(* Logix 5000 project; controller TFF vendor 1 type 14 code 107 rev 34.11; software revision 34.03; part 32 of 36 *)
(* tags used below, declared in another part *)
   FlowPathControl : FlowPathControl;   // Flow Path Control
   Options : Options;   // Options List
   PCV001_Control : PCV_Control;   // PCV001 Control UDT
   PCV101_Control : PCV_Control;   // PCV101 Control UDT
   PipeAnimation : PipeAnimation;   // HMI Pipe Animation Array
   XV001 : ALIAS FOR Valve[0];   // XV001
   XV002 : ALIAS FOR Valve[1];   // XV002
   XV004 : ALIAS FOR Valve[3];   // XV004
   XV005 : ALIAS FOR Valve[4];   // XV005
   XV006 : ALIAS FOR Valve[19];
   XV007 : ALIAS FOR Valve[20];
   XV102 : ALIAS FOR Valve[5];   // XV102
   XV401 : ALIAS FOR Valve[6];   // XV401
   XV402 : ALIAS FOR Valve[7];   // XV402
   XV403 : ALIAS FOR Valve[15];
   XV404 : ALIAS FOR Valve[16];
   XV405 : ALIAS FOR Valve[17];
   XV406 : ALIAS FOR Valve[18];
   XV411 : ALIAS FOR Valve[8];   // XV411
   XV421 : ALIAS FOR Valve[9];   // XV421
   XV431 : ALIAS FOR Valve[10];   // XV431
   XV441 : ALIAS FOR Valve[11];   // XV441
   XV501 : ALIAS FOR Valve[12];   // XV501
   XV502 : ALIAS FOR Valve[13];   // XV502
(* Process, continued *)

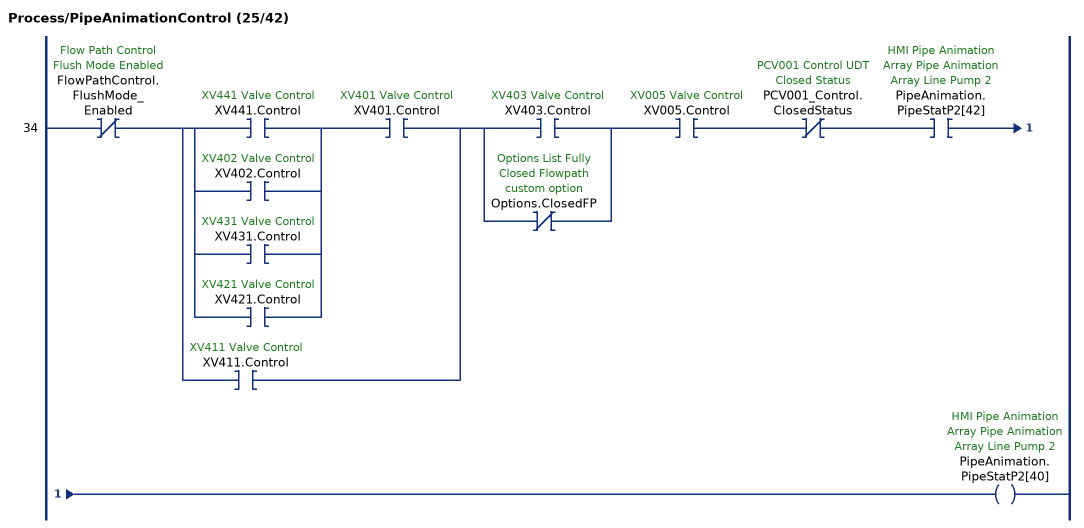
   [picture p389: Process/PipeAnimationControl rungs 34-34]
   34: XIO(FlowPathControl.FlushMode_Enabled)[[XIC(XV441.Control) ,XIC(XV402.Control) ,XIC(XV431.Control) ,XIC(XV421.Control) ] XIC(XV401.Control) ,XIC(XV411.Control) ][XIC(XV403.Control) ,XIO(Options.ClosedFP) ]XIC(XV005.Control)XIO(PCV001_Control.ClosedStatus)XIC(PipeAnimation.PipeStatP2[42])OTE(PipeAnimation.PipeStatP2[40]);
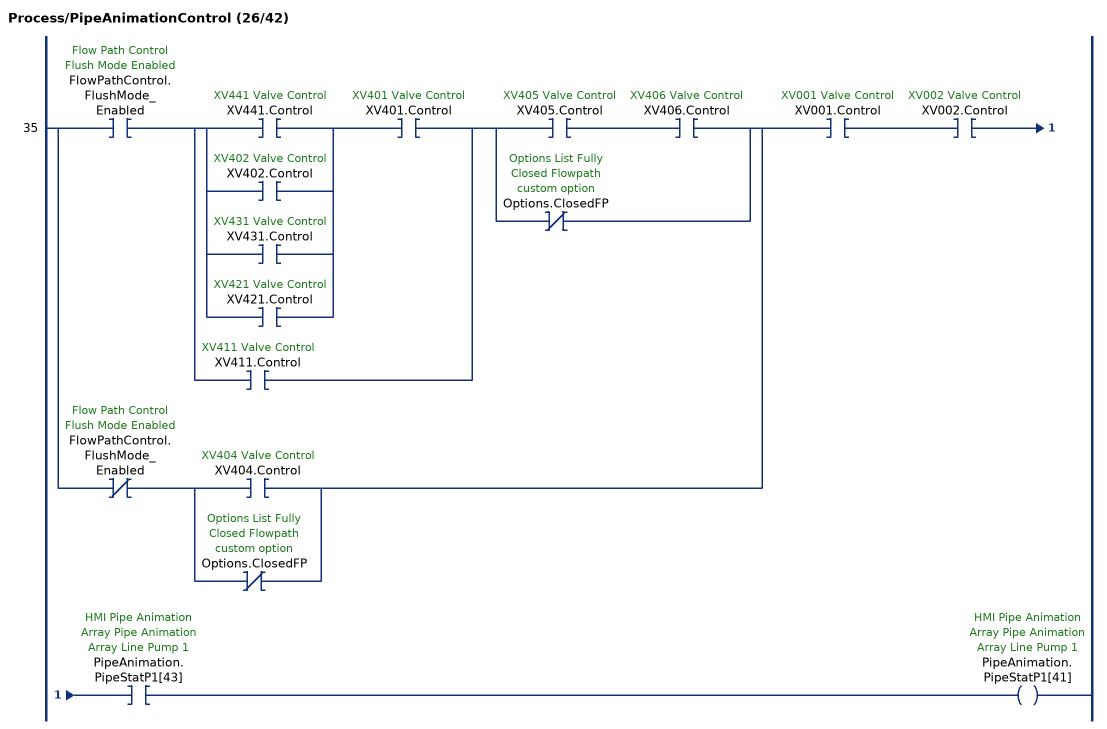
   35: [XIC(FlowPathControl.FlushMode_Enabled) [[XIC(XV441.Control) ,XIC(XV402.Control) ,XIC(XV431.Control) ,XIC(XV421.Control) ] XIC(XV401.Control) ,XIC(XV411.Control) ] [XIC(XV405.Control) XIC(XV406.Control) ,XIO(Options.ClosedFP) ] ,XIO(FlowPathControl.FlushMode_Enabled) [XIC(XV404.Control) ,XIO(Options.ClosedFP) ] ]XIC(XV001.Control)XIC(XV002.Control)XIC(PipeAnimation.PipeStatP1[43])OTE(PipeAnimation.PipeStatP1[41]);
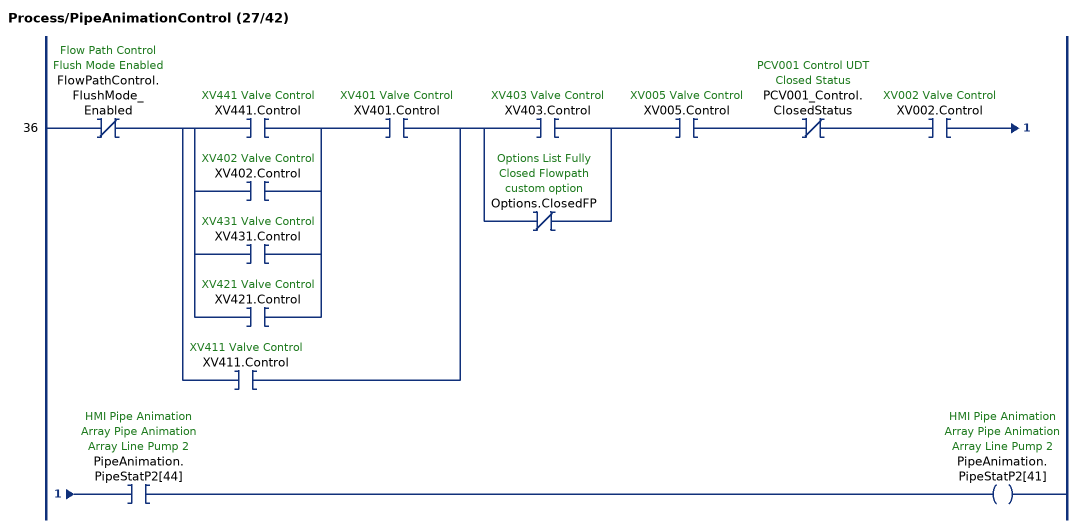
   36: XIO(FlowPathControl.FlushMode_Enabled)[[XIC(XV441.Control) ,XIC(XV402.Control) ,XIC(XV431.Control) ,XIC(XV421.Control) ] XIC(XV401.Control) ,XIC(XV411.Control) ][XIC(XV403.Control) ,XIO(Options.ClosedFP) ]XIC(XV005.Control)XIO(PCV001_Control.ClosedStatus)XIC(XV002.Control)XIC(PipeAnimation.PipeStatP2[44])OTE(PipeAnimation.PipeStatP2[41]);
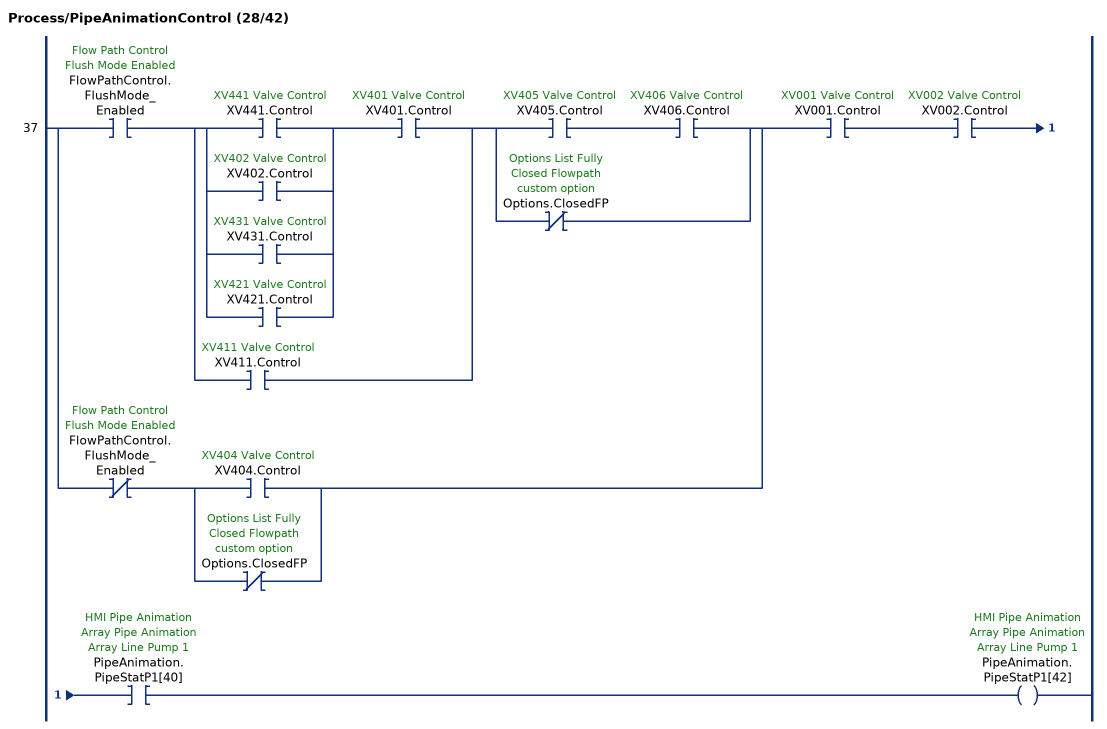
   37: [XIC(FlowPathControl.FlushMode_Enabled) [[XIC(XV441.Control) ,XIC(XV402.Control) ,XIC(XV431.Control) ,XIC(XV421.Control) ] XIC(XV401.Control) ,XIC(XV411.Control) ] [XIC(XV405.Control) XIC(XV406.Control) ,XIO(Options.ClosedFP) ] ,XIO(FlowPathControl.FlushMode_Enabled) [XIC(XV404.Control) ,XIO(Options.ClosedFP) ] ]XIC(XV001.Control)XIC(XV002.Control)XIC(PipeAnimation.PipeStatP1[40])OTE(PipeAnimation.PipeStatP1[42]);
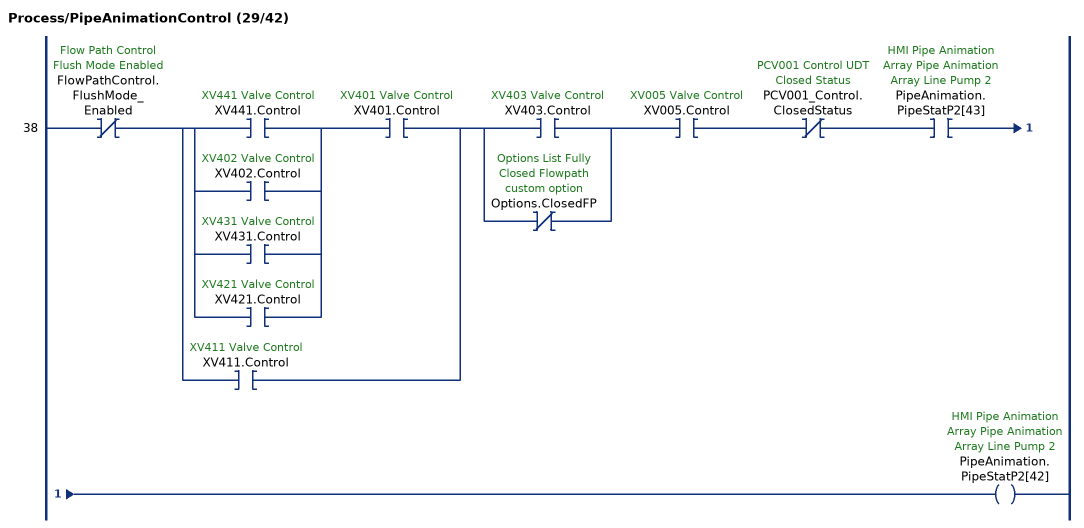
   38: XIO(FlowPathControl.FlushMode_Enabled)[[XIC(XV441.Control) ,XIC(XV402.Control) ,XIC(XV431.Control) ,XIC(XV421.Control) ] XIC(XV401.Control) ,XIC(XV411.Control) ][XIC(XV403.Control) ,XIO(Options.ClosedFP) ]XIC(XV005.Control)XIO(PCV001_Control.ClosedStatus)XIC(PipeAnimation.PipeStatP2[43])OTE(PipeAnimation.PipeStatP2[42]);
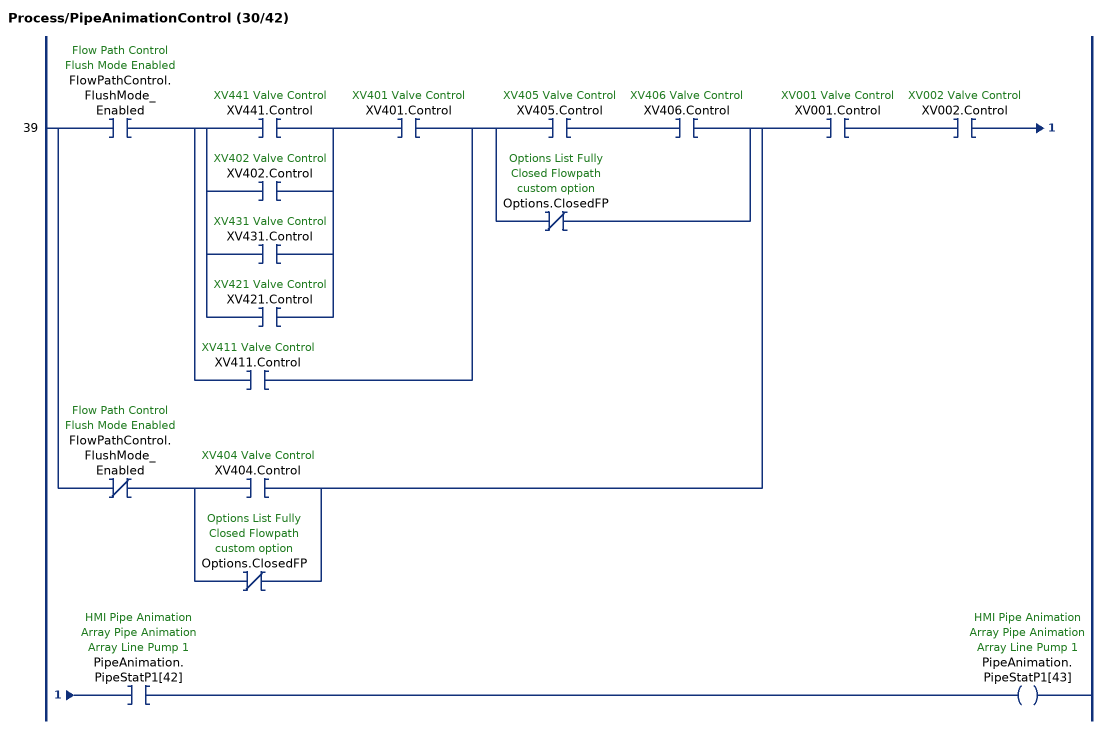
   39: [XIC(FlowPathControl.FlushMode_Enabled) [[XIC(XV441.Control) ,XIC(XV402.Control) ,XIC(XV431.Control) ,XIC(XV421.Control) ] XIC(XV401.Control) ,XIC(XV411.Control) ] [XIC(XV405.Control) XIC(XV406.Control) ,XIO(Options.ClosedFP) ] ,XIO(FlowPathControl.FlushMode_Enabled) [XIC(XV404.Control) ,XIO(Options.ClosedFP) ] ]XIC(XV001.Control)XIC(XV002.Control)XIC(PipeAnimation.PipeStatP1[42])OTE(PipeAnimation.PipeStatP1[43]);
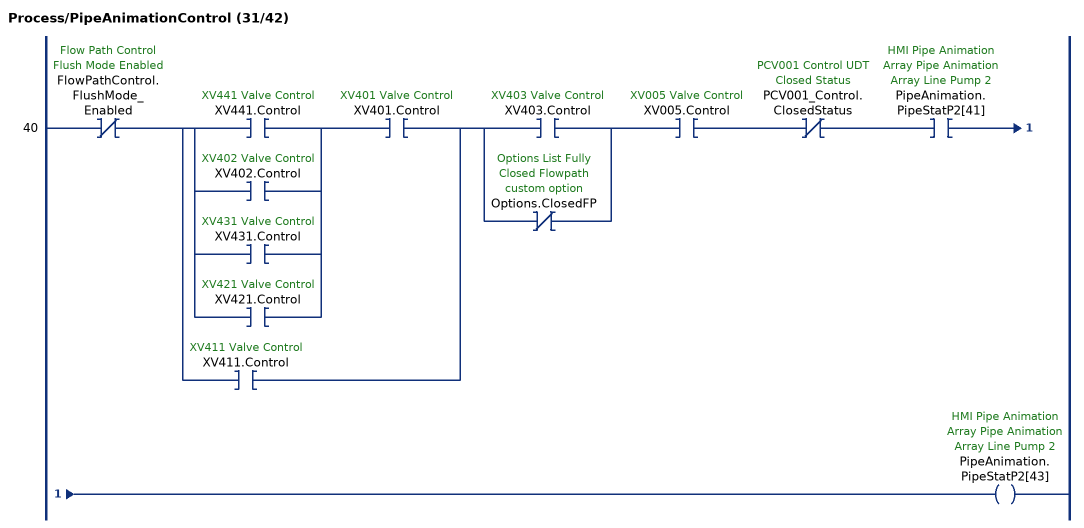
   40: XIO(FlowPathControl.FlushMode_Enabled)[[XIC(XV441.Control) ,XIC(XV402.Control) ,XIC(XV431.Control) ,XIC(XV421.Control) ] XIC(XV401.Control) ,XIC(XV411.Control) ][XIC(XV403.Control) ,XIO(Options.ClosedFP) ]XIC(XV005.Control)XIO(PCV001_Control.ClosedStatus)XIC(PipeAnimation.PipeStatP2[41])OTE(PipeAnimation.PipeStatP2[43]);
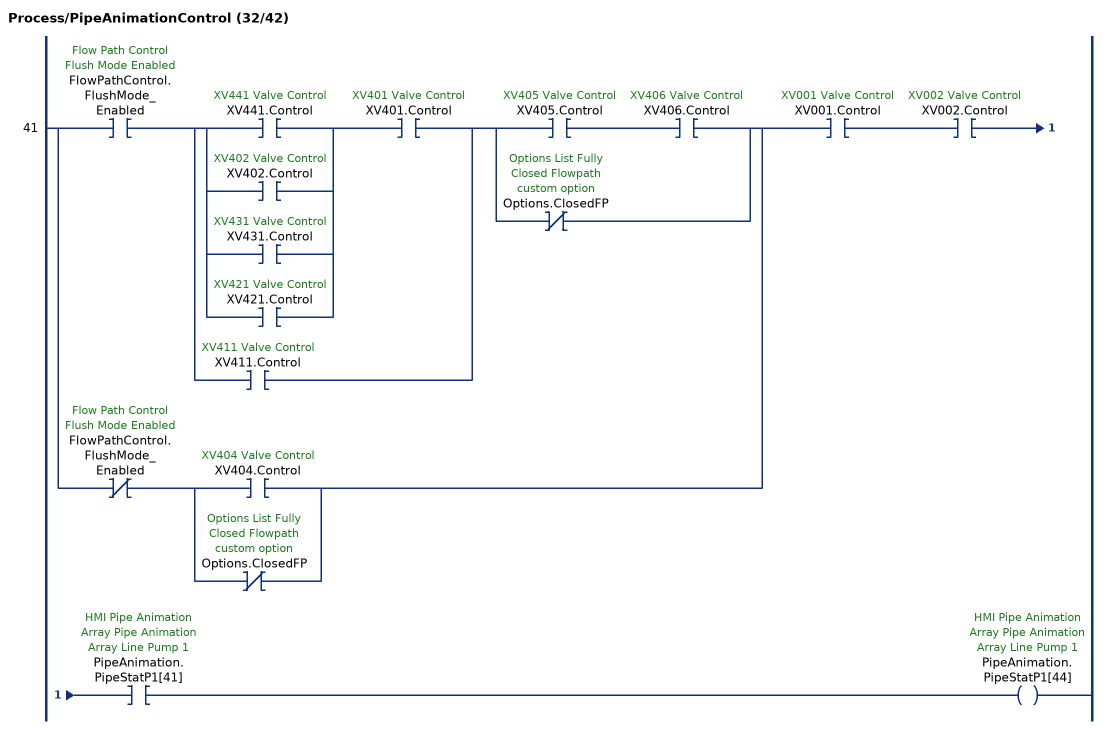
   41: [XIC(FlowPathControl.FlushMode_Enabled) [[XIC(XV441.Control) ,XIC(XV402.Control) ,XIC(XV431.Control) ,XIC(XV421.Control) ] XIC(XV401.Control) ,XIC(XV411.Control) ] [XIC(XV405.Control) XIC(XV406.Control) ,XIO(Options.ClosedFP) ] ,XIO(FlowPathControl.FlushMode_Enabled) [XIC(XV404.Control) ,XIO(Options.ClosedFP) ] ]XIC(XV001.Control)XIC(XV002.Control)XIC(PipeAnimation.PipeStatP1[41])OTE(PipeAnimation.PipeStatP1[44]);
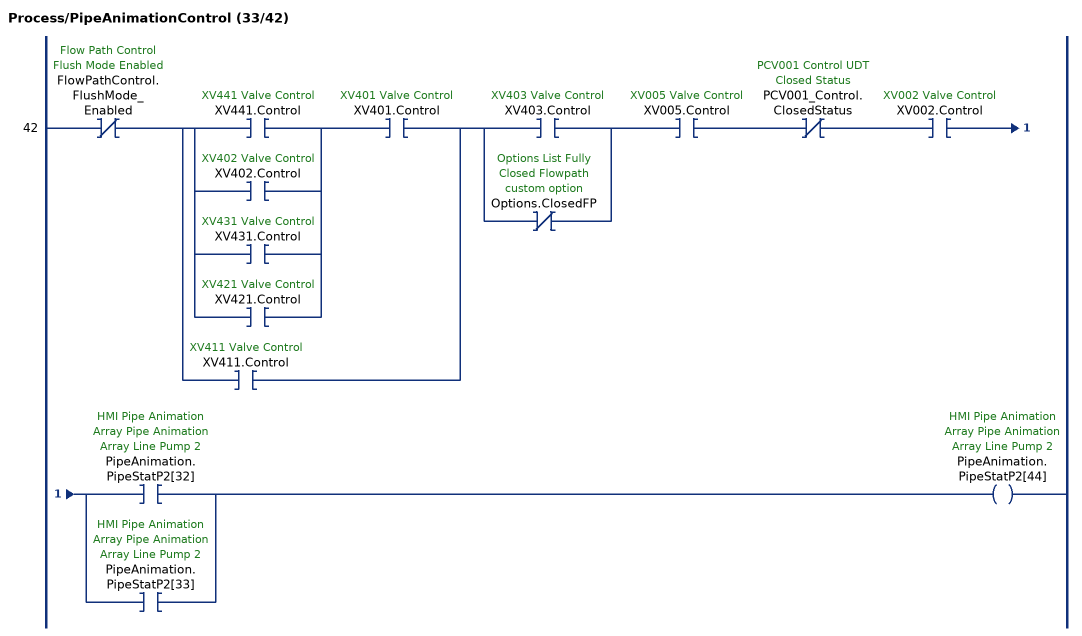
   42: XIO(FlowPathControl.FlushMode_Enabled)[[XIC(XV441.Control) ,XIC(XV402.Control) ,XIC(XV431.Control) ,XIC(XV421.Control) ] XIC(XV401.Control) ,XIC(XV411.Control) ][XIC(XV403.Control) ,XIO(Options.ClosedFP) ]XIC(XV005.Control)XIO(PCV001_Control.ClosedStatus)XIC(XV002.Control)[XIC(PipeAnimation.PipeStatP2[32]) ,XIC(PipeAnimation.PipeStatP2[33]) ]OTE(PipeAnimation.PipeStatP2[44]);
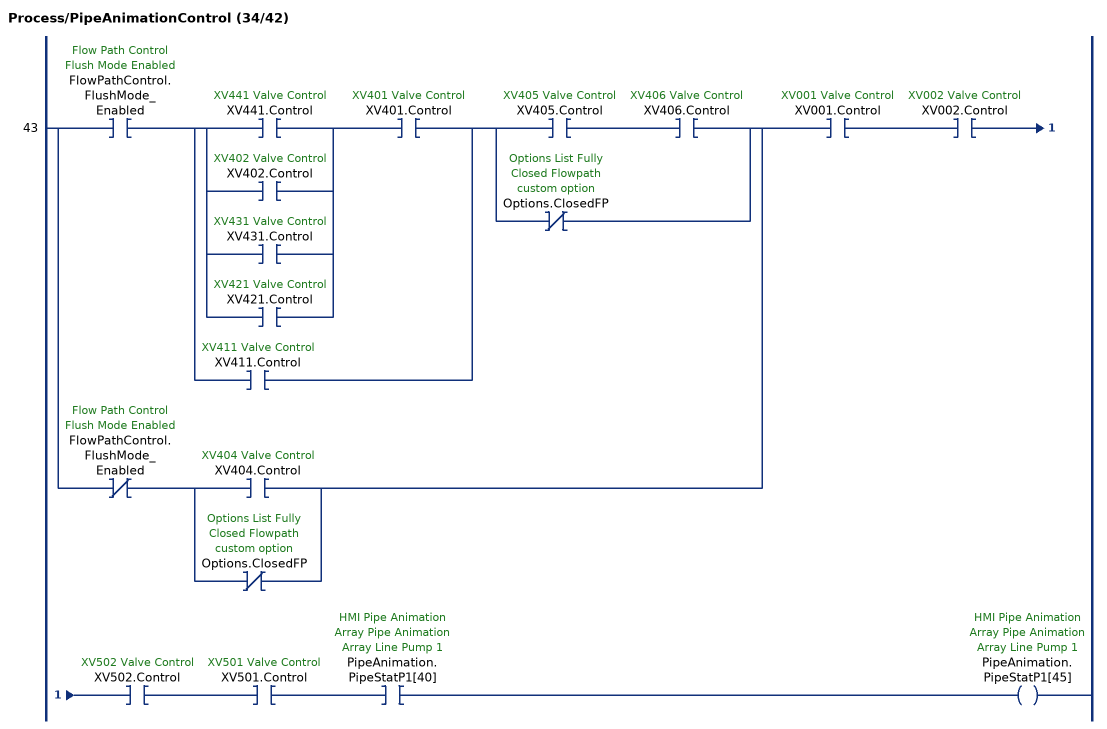
   43: [XIC(FlowPathControl.FlushMode_Enabled) [[XIC(XV441.Control) ,XIC(XV402.Control) ,XIC(XV431.Control) ,XIC(XV421.Control) ] XIC(XV401.Control) ,XIC(XV411.Control) ] [XIC(XV405.Control) XIC(XV406.Control) ,XIO(Options.ClosedFP) ] ,XIO(FlowPathControl.FlushMode_Enabled) [XIC(XV404.Control) ,XIO(Options.ClosedFP) ] ]XIC(XV001.Control)XIC(XV002.Control)XIC(XV502.Control)XIC(XV501.Control)XIC(PipeAnimation.PipeStatP1[40])OTE(PipeAnimation.PipeStatP1[45]);
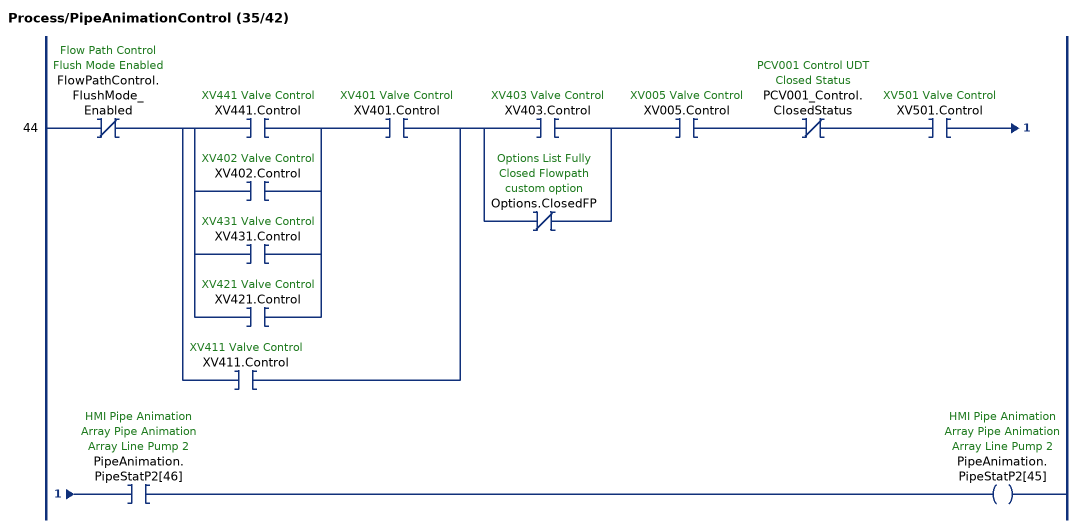
   44: XIO(FlowPathControl.FlushMode_Enabled)[[XIC(XV441.Control) ,XIC(XV402.Control) ,XIC(XV431.Control) ,XIC(XV421.Control) ] XIC(XV401.Control) ,XIC(XV411.Control) ][XIC(XV403.Control) ,XIO(Options.ClosedFP) ]XIC(XV005.Control)XIO(PCV001_Control.ClosedStatus)XIC(XV501.Control)XIC(PipeAnimation.PipeStatP2[46])OTE(PipeAnimation.PipeStatP2[45]);
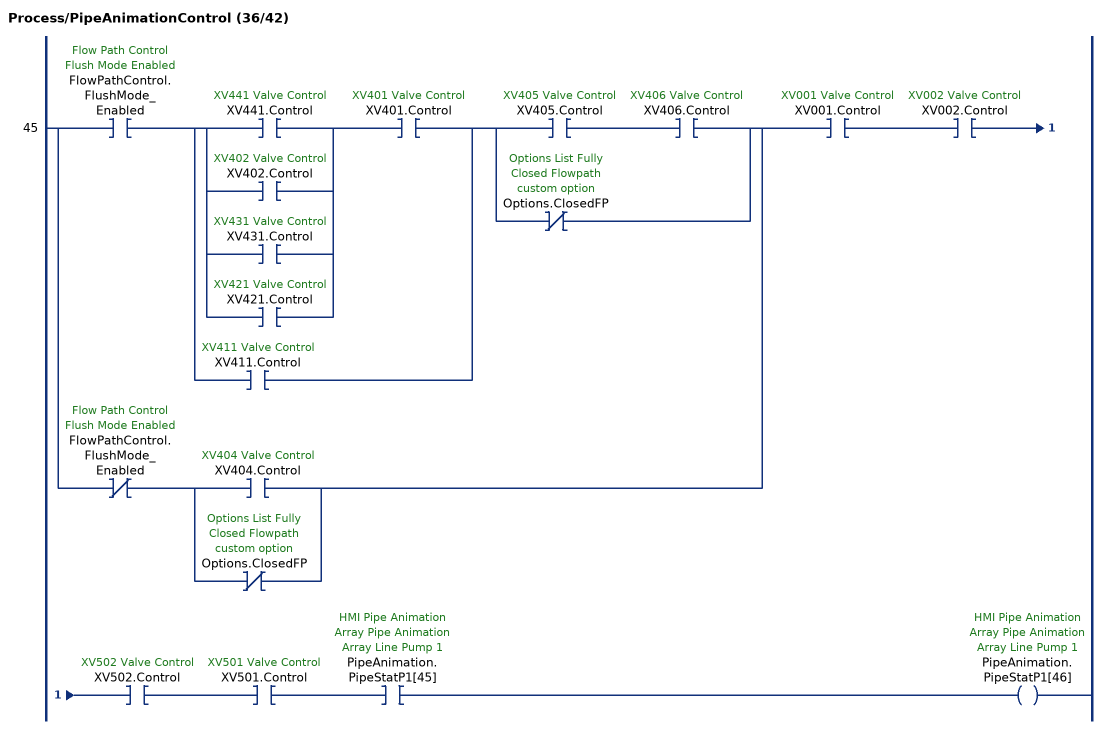
   45: [XIC(FlowPathControl.FlushMode_Enabled) [[XIC(XV441.Control) ,XIC(XV402.Control) ,XIC(XV431.Control) ,XIC(XV421.Control) ] XIC(XV401.Control) ,XIC(XV411.Control) ] [XIC(XV405.Control) XIC(XV406.Control) ,XIO(Options.ClosedFP) ] ,XIO(FlowPathControl.FlushMode_Enabled) [XIC(XV404.Control) ,XIO(Options.ClosedFP) ] ]XIC(XV001.Control)XIC(XV002.Control)XIC(XV502.Control)XIC(XV501.Control)XIC(PipeAnimation.PipeStatP1[45])OTE(PipeAnimation.PipeStatP1[46]);
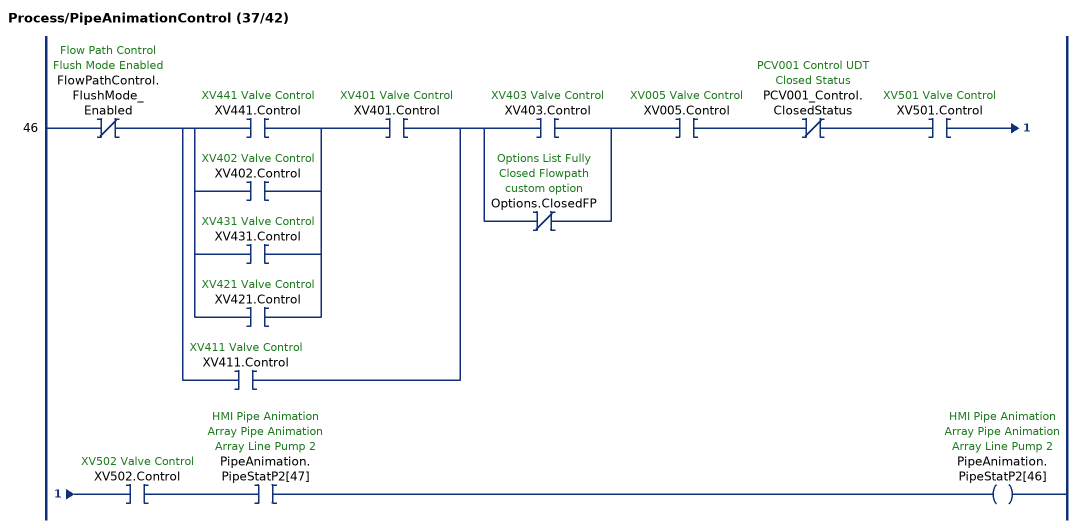
   46: XIO(FlowPathControl.FlushMode_Enabled)[[XIC(XV441.Control) ,XIC(XV402.Control) ,XIC(XV431.Control) ,XIC(XV421.Control) ] XIC(XV401.Control) ,XIC(XV411.Control) ][XIC(XV403.Control) ,XIO(Options.ClosedFP) ]XIC(XV005.Control)XIO(PCV001_Control.ClosedStatus)XIC(XV501.Control)XIC(XV502.Control)XIC(PipeAnimation.PipeStatP2[47])OTE(PipeAnimation.PipeStatP2[46]);
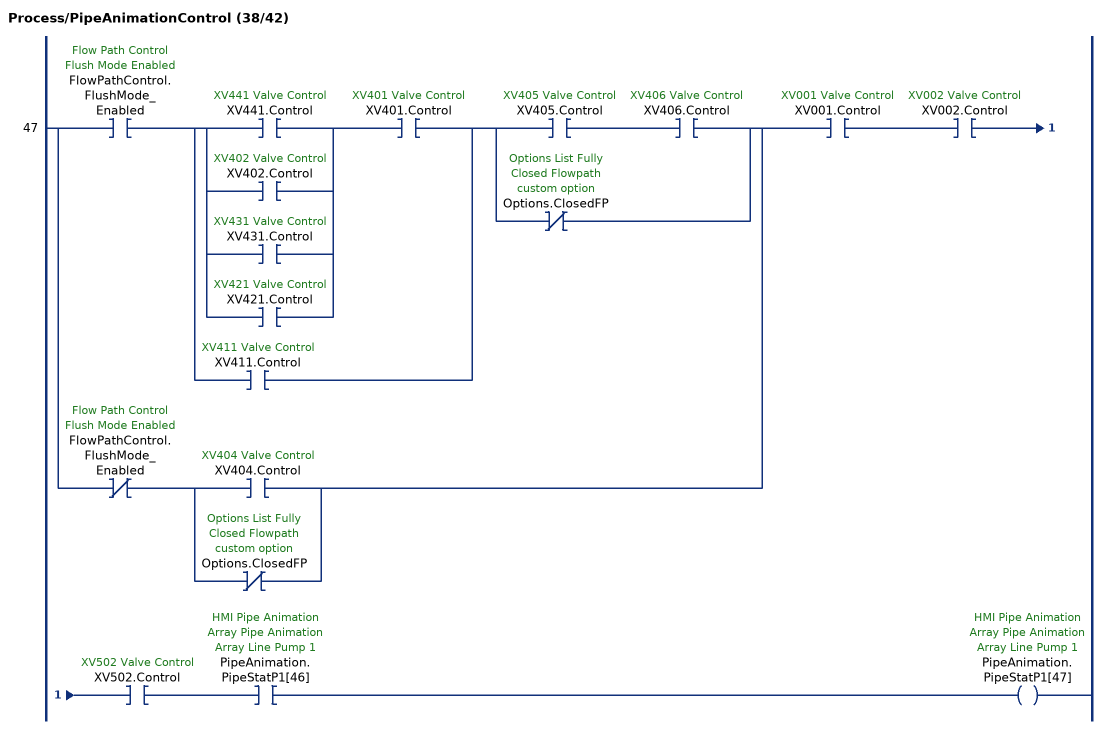
   47: [XIC(FlowPathControl.FlushMode_Enabled) [[XIC(XV441.Control) ,XIC(XV402.Control) ,XIC(XV431.Control) ,XIC(XV421.Control) ] XIC(XV401.Control) ,XIC(XV411.Control) ] [XIC(XV405.Control) XIC(XV406.Control) ,XIO(Options.ClosedFP) ] ,XIO(FlowPathControl.FlushMode_Enabled) [XIC(XV404.Control) ,XIO(Options.ClosedFP) ] ]XIC(XV001.Control)XIC(XV002.Control)XIC(XV502.Control)XIC(PipeAnimation.PipeStatP1[46])OTE(PipeAnimation.PipeStatP1[47]);
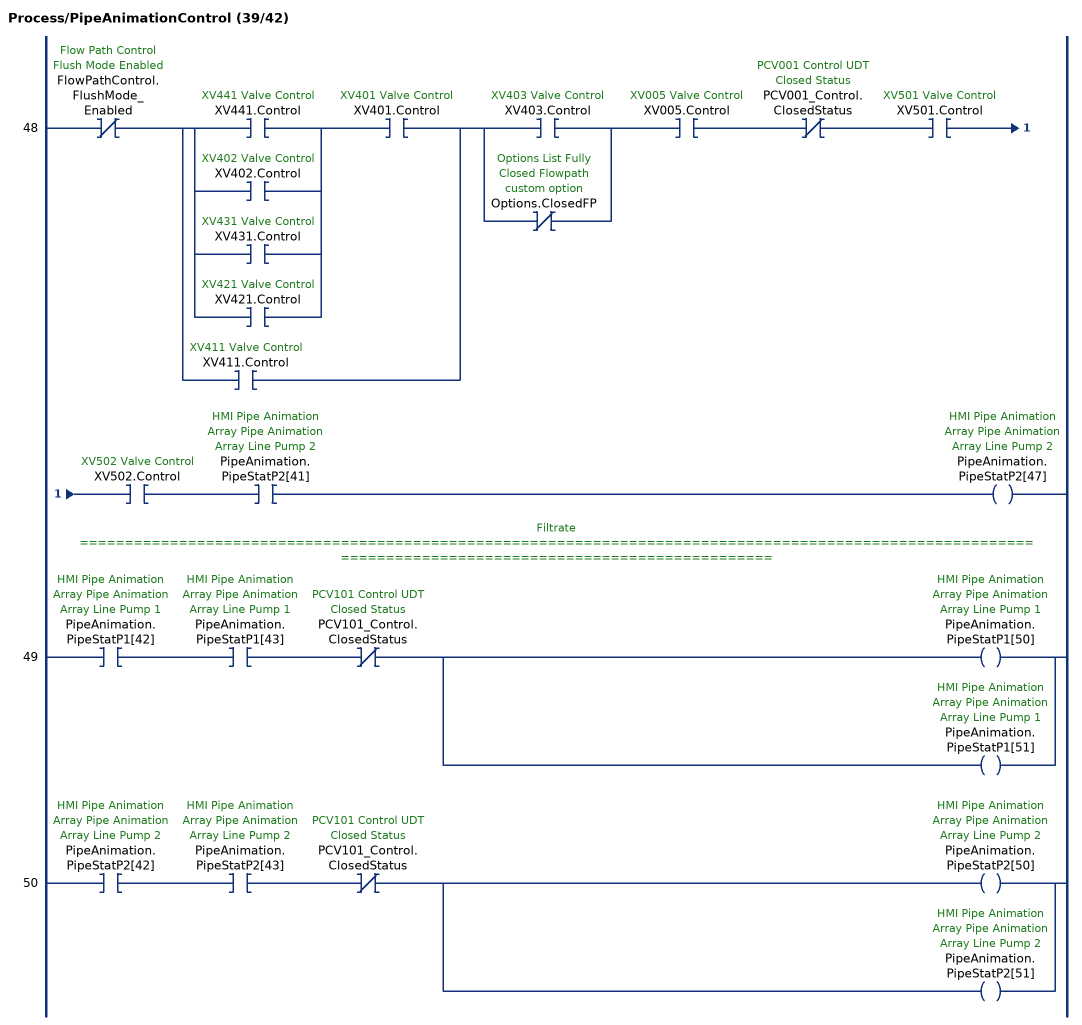
   48: XIO(FlowPathControl.FlushMode_Enabled)[[XIC(XV441.Control) ,XIC(XV402.Control) ,XIC(XV431.Control) ,XIC(XV421.Control) ] XIC(XV401.Control) ,XIC(XV411.Control) ][XIC(XV403.Control) ,XIO(Options.ClosedFP) ]XIC(XV005.Control)XIO(PCV001_Control.ClosedStatus)XIC(XV501.Control)XIC(XV502.Control)XIC(PipeAnimation.PipeStatP2[41])OTE(PipeAnimation.PipeStatP2[47]);
   // Filtrate
   // ==========================================================================================================================================================
   49: XIC(PipeAnimation.PipeStatP1[42])XIC(PipeAnimation.PipeStatP1[43])XIO(PCV101_Control.ClosedStatus)[OTE(PipeAnimation.PipeStatP1[50]) ,OTE(PipeAnimation.PipeStatP1[51]) ];
   50: XIC(PipeAnimation.PipeStatP2[42])XIC(PipeAnimation.PipeStatP2[43])XIO(PCV101_Control.ClosedStatus)[OTE(PipeAnimation.PipeStatP2[50]) ,OTE(PipeAnimation.PipeStatP2[51]) ];
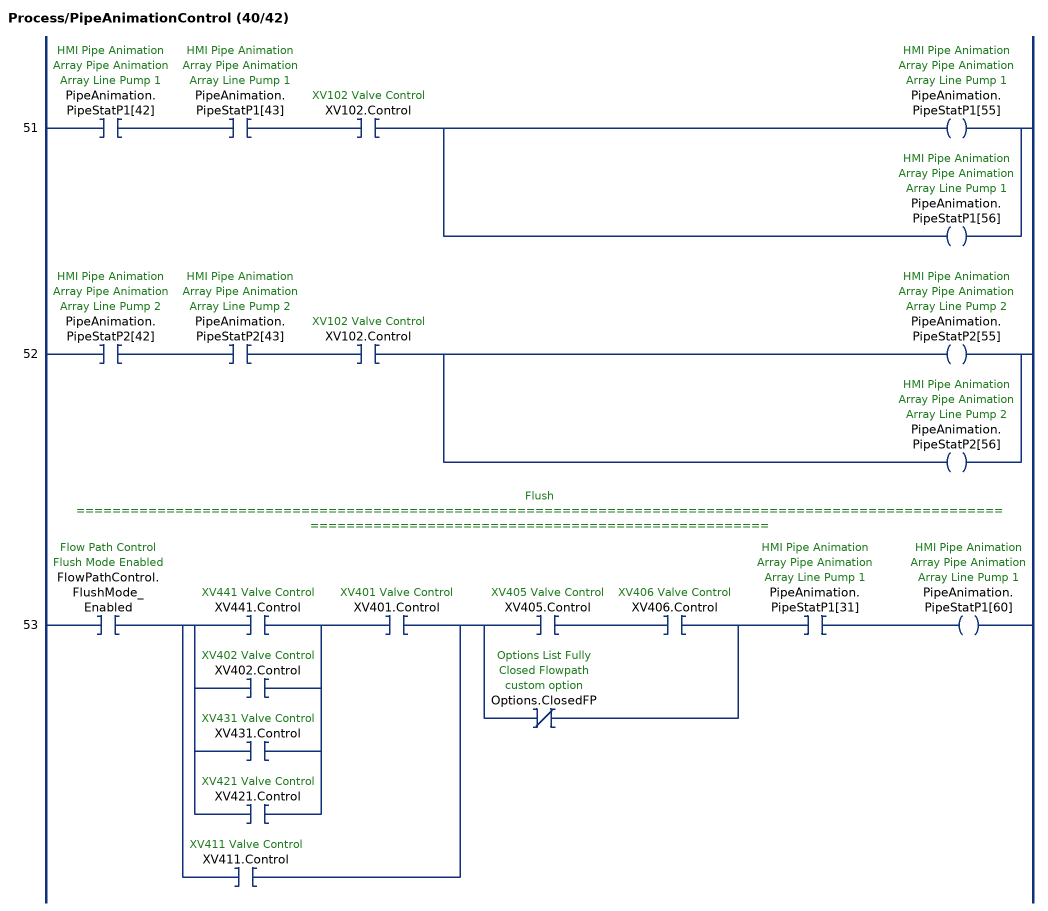
   51: XIC(PipeAnimation.PipeStatP1[42])XIC(PipeAnimation.PipeStatP1[43])XIC(XV102.Control)[OTE(PipeAnimation.PipeStatP1[55]) ,OTE(PipeAnimation.PipeStatP1[56]) ];
   52: XIC(PipeAnimation.PipeStatP2[42])XIC(PipeAnimation.PipeStatP2[43])XIC(XV102.Control)[OTE(PipeAnimation.PipeStatP2[55]) ,OTE(PipeAnimation.PipeStatP2[56]) ];
   // Flush
   // ==========================================================================================================================================================
   53: XIC(FlowPathControl.FlushMode_Enabled)[[XIC(XV441.Control) ,XIC(XV402.Control) ,XIC(XV431.Control) ,XIC(XV421.Control) ] XIC(XV401.Control) ,XIC(XV411.Control) ][XIC(XV405.Control) XIC(XV406.Control) ,XIO(Options.ClosedFP) ]XIC(PipeAnimation.PipeStatP1[31])OTE(PipeAnimation.PipeStatP1[60]);
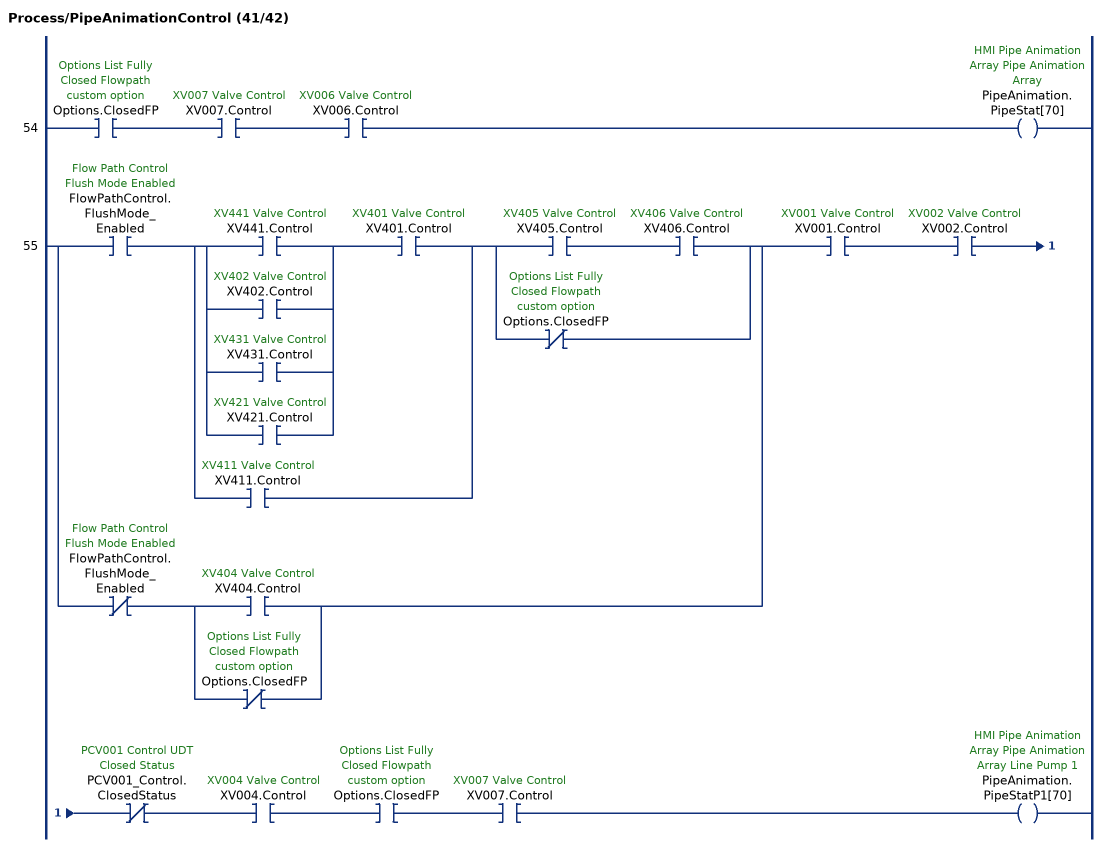
   54: XIC(Options.ClosedFP)XIC(XV007.Control)XIC(XV006.Control)OTE(PipeAnimation.PipeStat[70]);
   55: [XIC(FlowPathControl.FlushMode_Enabled) [[XIC(XV441.Control) ,XIC(XV402.Control) ,XIC(XV431.Control) ,XIC(XV421.Control) ] XIC(XV401.Control) ,XIC(XV411.Control) ] [XIC(XV405.Control) XIC(XV406.Control) ,XIO(Options.ClosedFP) ] ,XIO(FlowPathControl.FlushMode_Enabled) [XIC(XV404.Control) ,XIO(Options.ClosedFP) ] ]XIC(XV001.Control)XIC(XV002.Control)XIO(PCV001_Control.ClosedStatus)XIC(XV004.Control)XIC(Options.ClosedFP)XIC(XV007.Control)OTE(PipeAnimation.PipeStatP1[70]);
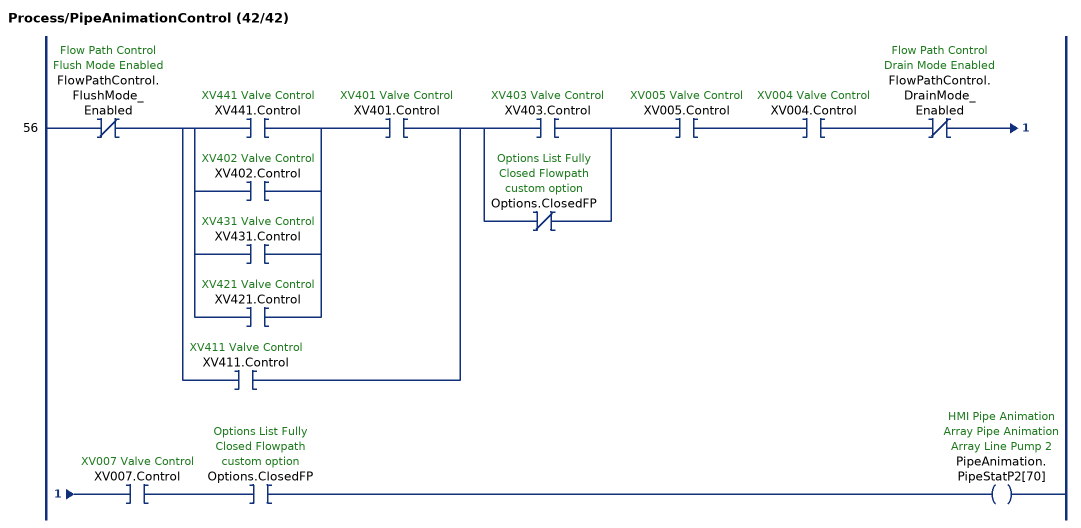
   56: XIO(FlowPathControl.FlushMode_Enabled)[[XIC(XV441.Control) ,XIC(XV402.Control) ,XIC(XV431.Control) ,XIC(XV421.Control) ] XIC(XV401.Control) ,XIC(XV411.Control) ][XIC(XV403.Control) ,XIO(Options.ClosedFP) ]XIC(XV005.Control)XIC(XV004.Control)XIO(FlowPathControl.DrainMode_Enabled)XIC(XV007.Control)XIC(Options.ClosedFP)OTE(PipeAnimation.PipeStatP2[70]);
END_ROUTINE
